Universal Robots URScript: T006_zai-org_GLM-4.7-FP8_edit_perf_rep1.urscript

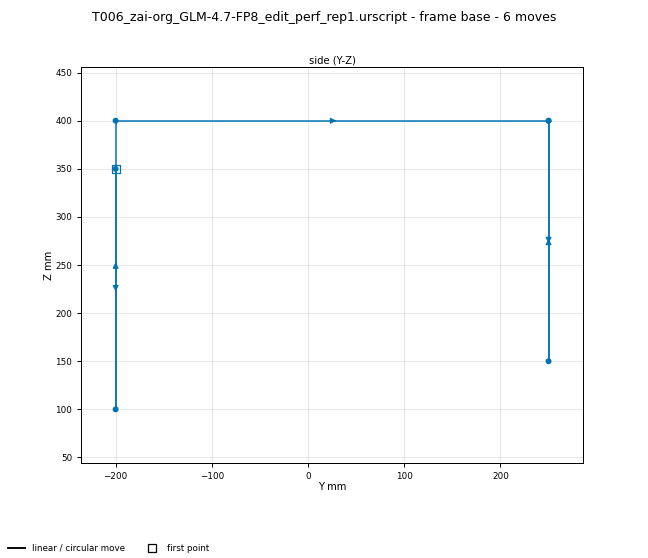
[picture p0: tool path of T006_zai-org_GLM-4.7-FP8_edit_perf_rep1.urscript in frame base, 6 of 8 moves have a stored position in this frame; points joined in program order, loops and branches not executed]
# Task: T006 — Bin picking with suction — fenced mode (Optimized)
# Generated by ENFIELD IR→URScript Translator
# Operating mode: fenced | Max TCP speed: 0.400 m/s
# Robot: ur5e
#
# WARNING: This is auto-generated code for SIMULATION ONLY.
# Do NOT deploy to a physical robot without safety review.

def task_T006():
  # [0] Verify E-Stop clear
  # E-Stop safety check (hardware-enforced on UR controller)
  if (get_digital_in(0) == True):
    popup("E-Stop active — aborting program.", error=True)
    halt
  end

  # [1] Home position
  # Optimized: Increased joint velocity and acceleration for faster transit
  movej([0.0000, -1.5708, 1.5708, -1.5708, -1.5708, 0.0000], a=2.5000, v=2.0000)

  # [2] Above bin
  # Optimized: Max TCP speed, increased acceleration, moderate blend
  movel(p[0.450000, -0.200000, 0.350000, 0.0000, 3.1416, 0.0000], a=2.5000, v=0.4000, r=0.0200)

  # [3] Descend into bin
  # Optimized: Increased approach speed, no blend for precision
  movel(p[0.450000, -0.200000, 0.100000, 0.0000, 3.1416, 0.0000], a=1.5000, v=0.2500)

  # [4] Suction ON
  set_digital_out(0, True)

  # [5] Vacuum settle
  # Optimized: Reduced settle time for faster cycle
  sleep(0.2000)

  # [6] Lift from bin
  # Optimized: Max TCP speed, increased acceleration, larger blend for smooth cornering
  movel(p[0.450000, -0.200000, 0.400000, 0.0000, 3.1416, 0.0000], a=2.5000, v=0.4000, r=0.0500)

  # [7] Transit to conveyor
  # Optimized: Max TCP speed, increased acceleration, larger blend
  movel(p[0.450000, 0.250000, 0.400000, 0.0000, 3.1416, 0.0000], a=2.5000, v=0.4000, r=0.0500)

  # [8] Descend to drop
  # Optimized: Increased drop speed, no blend for precision
  movel(p[0.450000, 0.250000, 0.150000, 0.0000, 3.1416, 0.0000], a=2.0000, v=0.3000)

  # [9] Suction OFF
  # Fixed: Corrected logic to False (OFF state)
  set_digital_out(0, False)

  # [10] Release settle
  # Optimized: Minimized wait time
  sleep(0.0500)

  # [11] Retract above conveyor
  # Optimized: Max TCP speed, increased acceleration, larger blend
  movel(p[0.450000, 0.250000, 0.400000, 0.0000, 3.1416, 0.0000], a=2.5000, v=0.4000, r=0.0500)

  # [12] Return to home
  # Optimized: Increased joint velocity and acceleration
  movej([0.0000, -1.5708, 1.5708, -1.5708, -1.5708, 0.0000], a=2.5000, v=2.0000)

end

# Entry point
task_T006()
